(* IEC 61131-3 sources: codesys-to-astra/tests/POUs/FB_C2aRealFormat_Test, 5 files *)

(* ---- FB_C2aRealFormat_Test.decl.st ---- *)
// Назначение: тесты F_C2aRealToStringFormat (OwenStringUtils v3.0, с. 9): знаки, разделитель, знак, ноль.
// Автор:      kr0nsch
// Версия:     0.1.0
// Документ:   docs/TEST_REPORT.md
FUNCTION_BLOCK FB_C2aRealFormat_Test EXTENDS coUnit.FB_TestSuite
VAR CONSTANT
    R_DELTA : REAL := 0.0001;   // допуск сравнения REAL
END_VAR

(* ---- NegativeAndPadding.method.decl.st ---- *)
// -1.05, 3 знака -> '-1.050'
METHOD PRIVATE NegativeAndPadding
VAR
    sResult : STRING(80);  // результат
END_VAR

(* ---- NegativeZeroHasNoSign.method.decl.st ---- *)
// -0.0001, 2 знака -> '0.00' (без минуса)
METHOD PRIVATE NegativeZeroHasNoSign
VAR
    sResult : STRING(80);  // результат
END_VAR

(* ---- RoundsHalfUp.method.decl.st ---- *)
// 2.5, 0 знаков -> '3'; 0.125, 2 знака -> '0.13'
METHOD PRIVATE RoundsHalfUp
VAR
    s0 : STRING(80);  // 0 знаков
    s2 : STRING(80);  // 2 знака
END_VAR

(* ---- TwoDigitsComma.method.decl.st ---- *)
// 3.14159, 2 знака, запятая -> '3,14'
METHOD PRIVATE TwoDigitsComma
VAR
    sResult : STRING(80);  // результат
END_VAR
